PROGRAM MAIN
VAR
	testall:testallfb;
END_VAR

testall();

END_PROGRAM

(* stored: Version 1.1.0.1, ProductVersion 3.1.4024.16
   POU MAIN: Id {d940760c-e873-4381-91d3-7b00ae51dd95}, SpecialFunc None *)
